(* IEC 61131-3 sources: plc-st-test/packages/core/test/testdata/interpreter, 24 files *)

(* ---- arrays.st ---- *)
(* IEC 61131-3 §6.4.4.4 / Table 15 (ARRAY): bounds are declared as [lo..hi] and may be negative or non-zero based; an element outside the declared bounds is a runtime error; arrays have value semantics on assignment (a copy, not an alias); multi-dimensional arrays index per dimension. *)
FUNCTION_BLOCK TEST_Arrays
VAR
  a : ARRAY[1..5] OF DINT;
  neg : ARRAY[-2..2] OF INT;
  m : ARRAY[0..1, 0..2] OF DINT;
  b : ARRAY[1..5] OF DINT;
  i, idx : DINT;
END_VAR
METHOD Test_FirstAndLastElement
  a[1] := 10;
  a[5] := 50;
  ASSERT_EQUAL_DINT(a[1], 10);
  ASSERT_EQUAL_DINT(a[5], 50);
  ASSERT_EQUAL_DINT(a[3], 0);
END_METHOD
METHOD Test_NegativeLowerBound
  neg[-2] := -20;
  neg[0] := 5;
  neg[2] := 22;
  ASSERT_EQUAL_INT(neg[-2], -20);
  ASSERT_EQUAL_INT(neg[0], 5);
  ASSERT_EQUAL_INT(neg[2], 22);
END_METHOD
METHOD Test_IndexBelowLowerBoundErrors
  idx := 0;
  a[idx] := 1;
END_METHOD
METHOD Test_IndexAboveUpperBoundErrors
  idx := 6;
  i := a[idx];
END_METHOD
METHOD Test_TwoDimensional
  FOR i := 0 TO 2 DO
    m[0, i] := i;
    m[1, i] := 10 + i;
  END_FOR
  ASSERT_EQUAL_DINT(m[0, 2], 2);
  ASSERT_EQUAL_DINT(m[1, 0], 10);
  ASSERT_EQUAL_DINT(m[1, 2], 12);
END_METHOD
METHOD Test_AssignmentCopiesValue
  a[1] := 1; a[2] := 2;
  b := a;
  a[1] := 99;
  ASSERT_EQUAL_DINT(b[1], 1);
  ASSERT_EQUAL_DINT(b[2], 2);
  ASSERT_EQUAL_DINT(a[1], 99);
END_METHOD
METHOD Test_ComputedIndex
  FOR i := 1 TO 5 DO
    a[i] := i * i;
  END_FOR
  ASSERT_EQUAL_DINT(a[a[2]], 16);
END_METHOD
END_FUNCTION_BLOCK

(* ---- bit-operations.st ---- *)
(* IEC 61131-3 §6.6.1 / Table 30 and Table 33: AND/OR/XOR/NOT on bit-string types work bitwise within the type's width (NOT BYTE#16#0F is 16#F0, not a wider value), and BOOL operands use plain logic. *)
FUNCTION_BLOCK TEST_BitOperations
VAR b : BYTE; w : WORD; dw : DWORD; lw : LWORD; END_VAR
METHOD Test_NotStaysInWidth
  b := 16#0F;
  ASSERT_EQUAL_BYTE(NOT b, 16#F0);
  w := 16#00FF;
  ASSERT_EQUAL_WORD(NOT w, 16#FF00);
  dw := 0;
  ASSERT_EQUAL_DWORD(NOT dw, 16#FFFFFFFF);
END_METHOD
METHOD Test_AndOrXor
  b := 16#CC;
  ASSERT_EQUAL_BYTE(b AND 16#0F, 16#0C);
  ASSERT_EQUAL_BYTE(b OR 16#0F, 16#CF);
  ASSERT_EQUAL_BYTE(b XOR 16#FF, 16#33);
END_METHOD
METHOD Test_WordMasks
  w := 16#ABCD;
  ASSERT_EQUAL_WORD(w AND 16#FF00, 16#AB00);
  ASSERT_EQUAL_WORD(w AND 16#00FF, 16#00CD);
  ASSERT_EQUAL_WORD(w XOR w, 0);
END_METHOD
METHOD Test_Lword64BitOps
  lw := 16#8000_0000_0000_0001;
  ASSERT_EQUAL_LWORD(lw AND 16#FFFF_FFFF_0000_0000, 16#8000_0000_0000_0000);
  ASSERT_EQUAL_LWORD(lw OR 16#2, 16#8000_0000_0000_0003);
  ASSERT_EQUAL_LWORD(NOT lw, 16#7FFF_FFFF_FFFF_FFFE);
END_METHOD
METHOD Test_BoolLogicTruthTables
  ASSERT_TRUE(TRUE AND TRUE);
  ASSERT_FALSE(TRUE AND FALSE);
  ASSERT_TRUE(FALSE OR TRUE);
  ASSERT_FALSE(FALSE OR FALSE);
  ASSERT_FALSE(TRUE XOR TRUE);
  ASSERT_TRUE(TRUE XOR FALSE);
  ASSERT_TRUE(NOT FALSE);
  ASSERT_FALSE(NOT TRUE);
END_METHOD
END_FUNCTION_BLOCK

(* ---- case-statement.st ---- *)
(* IEC 61131-3 §6.6.2.5.3 / Table 72 (CASE): selector arms may be single values, comma lists and ranges a..b; ELSE runs when no arm matches; at most one arm runs; enumerated selectors use enumerator labels. *)
TYPE E_Mode : (Off, Manual, Auto, Fault); END_TYPE

FUNCTION_BLOCK TEST_Case
VAR n, r : DINT; m : E_Mode; END_VAR
METHOD Classify
  CASE n OF
    1: r := 10;
    2, 3, 5: r := 20;
    10..19: r := 30;
    -5..-1: r := 40;
  ELSE
    r := 99;
  END_CASE
END_METHOD
METHOD Test_SingleValue
  n := 1; Classify();
  ASSERT_EQUAL_DINT(r, 10);
END_METHOD
METHOD Test_List
  n := 2; Classify();
  ASSERT_EQUAL_DINT(r, 20);
  n := 3; Classify();
  ASSERT_EQUAL_DINT(r, 20);
  n := 5; Classify();
  ASSERT_EQUAL_DINT(r, 20);
END_METHOD
METHOD Test_ListGapFallsToElse
  n := 4; Classify();
  ASSERT_EQUAL_DINT(r, 99);
END_METHOD
METHOD Test_RangeBounds
  n := 10; Classify();
  ASSERT_EQUAL_DINT(r, 30);
  n := 15; Classify();
  ASSERT_EQUAL_DINT(r, 30);
  n := 19; Classify();
  ASSERT_EQUAL_DINT(r, 30);
  n := 9; Classify();
  ASSERT_EQUAL_DINT(r, 99);
  n := 20; Classify();
  ASSERT_EQUAL_DINT(r, 99);
END_METHOD
METHOD Test_NegativeRange
  n := -3; Classify();
  ASSERT_EQUAL_DINT(r, 40);
  n := 0; Classify();
  ASSERT_EQUAL_DINT(r, 99);
END_METHOD
METHOD Test_NoElseNoMatchLeavesUnchanged
  r := 7; n := 50;
  CASE n OF
    1: r := 1;
  END_CASE
  ASSERT_EQUAL_DINT(r, 7);
END_METHOD
METHOD Test_EnumArms
  m := E_Mode.Auto;
  CASE m OF
    E_Mode.Off: r := 0;
    E_Mode.Manual, E_Mode.Auto: r := 1;
    E_Mode.Fault: r := 2;
  END_CASE
  ASSERT_EQUAL_DINT(r, 1);
  m := E_Mode.Fault;
  CASE m OF
    E_Mode.Off: r := 0;
    E_Mode.Manual, E_Mode.Auto: r := 1;
    E_Mode.Fault: r := 2;
  END_CASE
  ASSERT_EQUAL_DINT(r, 2);
END_METHOD
METHOD Test_EnumElse
  m := E_Mode.Manual;
  CASE m OF
    E_Mode.Off: r := 0;
  ELSE
    r := -1;
  END_CASE
  ASSERT_EQUAL_DINT(r, -1);
END_METHOD
METHOD Test_OnlyFirstMatchingArmRuns
  n := 2; r := 0;
  CASE n OF
    1..5: r := r + 1;
    2: r := r + 100;
  END_CASE
  ASSERT_EQUAL_DINT(r, 1);
END_METHOD
END_FUNCTION_BLOCK

(* ---- conversions.st ---- *)
(* IEC 61131-3 §6.6.1 Table 30 note on conversion: REAL/LREAL to an integer type rounds to nearest, ties to even (so 0.5 -> 0, 1.5 -> 2, 2.5 -> 2, -0.5 -> 0, -1.5 -> -2); integer narrowing keeps the low-order bits (two's complement wrap); BOOL converts to 0/1. *)
FUNCTION_BLOCK TEST_Conversions
VAR r : REAL; l : LREAL; i : INT; d : DINT; END_VAR
METHOD Test_RealToIntTiesToEven
  r := 0.5;
  ASSERT_EQUAL_DINT(REAL_TO_DINT(r), 0);
  r := 1.5;
  ASSERT_EQUAL_DINT(REAL_TO_DINT(r), 2);
  r := 2.5;
  ASSERT_EQUAL_DINT(REAL_TO_DINT(r), 2);
  r := 3.5;
  ASSERT_EQUAL_DINT(REAL_TO_DINT(r), 4);
END_METHOD
METHOD Test_NegativeTiesToEven
  r := -0.5;
  ASSERT_EQUAL_DINT(REAL_TO_DINT(r), 0);
  r := -1.5;
  ASSERT_EQUAL_DINT(REAL_TO_DINT(r), -2);
  r := -2.5;
  ASSERT_EQUAL_DINT(REAL_TO_DINT(r), -2);
END_METHOD
METHOD Test_NonTiesRoundToNearest
  l := 2.4;
  ASSERT_EQUAL_DINT(LREAL_TO_DINT(l), 2);
  l := 2.6;
  ASSERT_EQUAL_DINT(LREAL_TO_DINT(l), 3);
  l := -2.6;
  ASSERT_EQUAL_DINT(LREAL_TO_DINT(l), -3);
END_METHOD
METHOD Test_IntNarrowingWraps
  d := 300;
  ASSERT_EQUAL_SINT(DINT_TO_SINT(d), 44);
  d := 70000;
  ASSERT_EQUAL_INT(DINT_TO_INT(d), 4464);
  d := -1;
  ASSERT_EQUAL_USINT(DINT_TO_USINT(d), 255);
END_METHOD
METHOD Test_WideningPreservesValue
  i := -5;
  ASSERT_EQUAL_DINT(INT_TO_DINT(i), -5);
  ASSERT_EQUAL_LINT(INT_TO_LINT(i), -5);
  ASSERT_EQUAL_REAL(INT_TO_REAL(i), -5.0);
END_METHOD
METHOD Test_BoolConversions
  ASSERT_EQUAL_DINT(BOOL_TO_DINT(TRUE), 1);
  ASSERT_EQUAL_DINT(BOOL_TO_DINT(FALSE), 0);
  d := 7;
  ASSERT_TRUE(DINT_TO_BOOL(d));
  d := 0;
  ASSERT_FALSE(DINT_TO_BOOL(d));
END_METHOD
METHOD Test_UnsignedFromNegativeWraps
  d := -1;
  ASSERT_EQUAL_UDINT(DINT_TO_UDINT(d), 4294967295);
END_METHOD
END_FUNCTION_BLOCK

(* ---- counters-edges.st ---- *)
(* IEC 61131-3 §6.6.3.2 / Tables 41-42 (CTU, CTD) and R_TRIG/F_TRIG (Table 40): counters count only on a rising edge of CU/CD evaluated once per cycle, so holding the input TRUE for many cycles counts once; CTU.Q = (CV >= PV); R_TRIG.Q is TRUE for exactly the cycle in which CLK rose. *)
FUNCTION_BLOCK TEST_CountersEdges
VAR
  ctu : CTU;
  rt : R_TRIG;
  ft : F_TRIG;
  clk : BOOL;
  rst : BOOL;
  rises, falls : DINT;
END_VAR
METHOD Cycle
  ctu(CU := clk, R := rst, PV := 3);
  rt(CLK := clk);
  ft(CLK := clk);
  IF rt.Q THEN rises := rises + 1; END_IF
  IF ft.Q THEN falls := falls + 1; END_IF
END_METHOD
METHOD Test_HeldInputCountsOnce
  clk := TRUE;
  RUN_CYCLES(10);
  ASSERT_EQUAL_INT(ctu.CV, 1);
  ASSERT_EQUAL_DINT(rises, 1);
  ASSERT_EQUAL_DINT(falls, 0);
END_METHOD
METHOD Test_ToggleCountsEachRisingEdge
  clk := TRUE;  RUN_CYCLES(1);
  clk := FALSE; RUN_CYCLES(1);
  clk := TRUE;  RUN_CYCLES(1);
  clk := FALSE; RUN_CYCLES(1);
  ASSERT_EQUAL_INT(ctu.CV, 2);
  ASSERT_EQUAL_DINT(rises, 2);
  ASSERT_EQUAL_DINT(falls, 2);
  ASSERT_FALSE(ctu.Q);
END_METHOD
METHOD Test_QSetsAtPreset
  clk := TRUE;  RUN_CYCLES(1);
  clk := FALSE; RUN_CYCLES(1);
  clk := TRUE;  RUN_CYCLES(1);
  clk := FALSE; RUN_CYCLES(1);
  clk := TRUE;  RUN_CYCLES(1);
  ASSERT_EQUAL_INT(ctu.CV, 3);
  ASSERT_TRUE(ctu.Q);
END_METHOD
METHOD Test_ResetClearsCountAndQ
  clk := TRUE;  RUN_CYCLES(1);
  clk := FALSE; RUN_CYCLES(1);
  clk := TRUE;  RUN_CYCLES(1);
  clk := FALSE; RUN_CYCLES(1);
  clk := TRUE;  RUN_CYCLES(1);
  rst := TRUE;
  RUN_CYCLES(1);
  ASSERT_EQUAL_INT(ctu.CV, 0);
  ASSERT_FALSE(ctu.Q);
END_METHOD
METHOD Test_PulseOnlyOneCycleWide
  clk := TRUE;
  RUN_CYCLES(1);
  ASSERT_TRUE(rt.Q);
  RUN_CYCLES(1);
  ASSERT_FALSE(rt.Q);
END_METHOD
END_FUNCTION_BLOCK

(* ---- deep-nesting.st ---- *)
(* IEC 61131-3 §6.6.2 (statements compose freely): IF/ELSIF/ELSE, CASE and loops nest to arbitrary depth with the innermost branch selected by the combined conditions; expressions nest through parentheses with the Table 71 precedence (NOT, **, unary minus, * / MOD, + -, comparisons, AND, XOR, OR). *)
FUNCTION_BLOCK TEST_DeepNesting
VAR a, b, c, r, i, j, k, count : DINT; ok : BOOL; END_VAR
METHOD Test_NestedIfElsifChain
  a := 2; b := 3; c := 4;
  IF a = 1 THEN
    r := 1;
  ELSIF a = 2 THEN
    IF b = 2 THEN
      r := 2;
    ELSIF b = 3 THEN
      IF c = 3 THEN
        r := 3;
      ELSE
        IF c = 4 THEN r := 4; ELSE r := 5; END_IF
      END_IF
    END_IF
  ELSE
    r := 6;
  END_IF
  ASSERT_EQUAL_DINT(r, 4);
END_METHOD
METHOD Test_TripleNestedLoopCount
  count := 0;
  FOR i := 1 TO 4 DO
    FOR j := 1 TO 3 DO
      FOR k := 1 TO 2 DO
        count := count + 1;
      END_FOR
    END_FOR
  END_FOR
  ASSERT_EQUAL_DINT(count, 24);
END_METHOD
METHOD Test_LoopsCaseAndIfTogether
  count := 0;
  FOR i := 1 TO 6 DO
    CASE i MOD 3 OF
      0: count := count + 100;
      1:
        IF i > 3 THEN count := count + 10; ELSE count := count + 1; END_IF
    ELSE
      count := count + 1000;
    END_CASE
  END_FOR
  ASSERT_EQUAL_DINT(count, 2 * 1000 + 2 * 100 + 10 + 1);
END_METHOD
METHOD Test_ParenthesesNestDeeply
  a := 2;
  r := ((((a + 1) * (a + 2)) - ((a - 1) * (a + 3))) * 2) + (((a)));
  ASSERT_EQUAL_DINT(r, 16);
END_METHOD
METHOD Test_PrecedenceTable71
  r := 2 + 3 * 4;
  ASSERT_EQUAL_DINT(r, 14);
  r := 20 - 6 / 3 - 1;
  ASSERT_EQUAL_DINT(r, 17);
  r := 2 * 3 MOD 4;
  ASSERT_EQUAL_DINT(r, 2);
  r := -2 * 3;
  ASSERT_EQUAL_DINT(r, -6);
END_METHOD
METHOD Test_BooleanPrecedence
  ok := TRUE OR FALSE AND FALSE;
  ASSERT_TRUE(ok);
  ok := NOT FALSE AND FALSE;
  ASSERT_FALSE(ok);
  ok := TRUE XOR TRUE OR TRUE;
  ASSERT_TRUE(ok);
  a := 1; b := 2;
  ok := a < b AND b < 3 OR FALSE;
  ASSERT_TRUE(ok);
END_METHOD
METHOD Test_WhileInsideRepeatInsideFor
  count := 0;
  FOR i := 1 TO 2 DO
    j := 0;
    REPEAT
      j := j + 1;
      k := 0;
      WHILE k < 2 DO
        k := k + 1;
        count := count + 1;
      END_WHILE
    UNTIL j >= 3
    END_REPEAT
  END_FOR
  ASSERT_EQUAL_DINT(count, 12);
END_METHOD
END_FUNCTION_BLOCK

(* ---- division.st ---- *)
(* IEC 61131-3 §6.6.1.4 / Table 30: division by zero is an error for integer and real operands, and for MOD; this runtime raises IecRuntimeError 'division by zero' (test errored). Also integer division truncates toward zero. *)
FUNCTION_BLOCK TEST_Division
VAR i, z : DINT; r, rz : REAL; l, lz : LREAL; END_VAR
METHOD Test_IntDivByZeroErrors
  z := 0; i := 5 / z;
END_METHOD
METHOD Test_RealDivByZeroErrors
  rz := 0.0; r := 1.0 / rz;
END_METHOD
METHOD Test_LrealDivByZeroErrors
  lz := 0.0; l := 1.0 / lz;
END_METHOD
METHOD Test_ModByZeroErrors
  z := 0; i := 5 MOD z;
END_METHOD
METHOD Test_IntDivTruncatesTowardZero
  i := 7; z := 2;
  ASSERT_EQUAL_DINT(i / z, 3);
  i := -7;
  ASSERT_EQUAL_DINT(i / z, -3);
  z := -2;
  ASSERT_EQUAL_DINT(i / z, 3);
  i := 7;
  ASSERT_EQUAL_DINT(i / z, -3);
END_METHOD
METHOD Test_RealDivNormal
  r := 1.0; rz := 4.0;
  ASSERT_EQUAL_REAL(r / rz, 0.25);
END_METHOD
END_FUNCTION_BLOCK

(* ---- enums.st ---- *)
(* IEC 61131-3 §6.4.4.2 / Table 12 (enumerated data types): enumerators without an explicit value number from 0 and continue from the previous value after an explicit one; a variable of enumerated type starts at its first enumerator unless an initial value is given; enumerators of one type compare by value. *)
TYPE E_Color : (Red, Green := 5, Blue); END_TYPE
TYPE E_Level : (Low, Mid, High) := Mid; END_TYPE

FUNCTION_BLOCK TEST_Enums
VAR
  c : E_Color;
  lv : E_Level;
  c2 : E_Color := E_Color.Blue;
  n : DINT;
END_VAR
METHOD Test_DefaultIsFirstEnumerator
  ASSERT_EQUAL(c, E_Color.Red);
END_METHOD
METHOD Test_DeclaredInitialValue
  ASSERT_EQUAL(c2, E_Color.Blue);
END_METHOD
METHOD Test_TypeLevelDefault
  ASSERT_EQUAL(lv, E_Level.Mid);
END_METHOD
METHOD Test_ExplicitAndImplicitValues
  n := E_Color.Red;
  ASSERT_EQUAL_DINT(n, 0);
  n := E_Color.Green;
  ASSERT_EQUAL_DINT(n, 5);
  n := E_Color.Blue;
  ASSERT_EQUAL_DINT(n, 6);
END_METHOD
METHOD Test_Comparison
  c := E_Color.Green;
  ASSERT_TRUE(c = E_Color.Green);
  ASSERT_TRUE(c <> E_Color.Blue);
  ASSERT_NOT_EQUAL(c, E_Color.Red);
END_METHOD
METHOD Test_AssignAndCopy
  c := E_Color.Blue;
  c2 := c;
  c := E_Color.Red;
  ASSERT_EQUAL(c2, E_Color.Blue);
  ASSERT_EQUAL(c, E_Color.Red);
END_METHOD
END_FUNCTION_BLOCK

(* ---- fb-instances.st ---- *)
(* IEC 61131-3 §6.6.3 (function blocks): every FB instance has its own copy of the internal VAR state, instances do not share data, and state persists between calls of the same instance. Struct assignment (§6.4.4.3) copies all members. *)
TYPE ST_Point : STRUCT x : DINT; y : DINT; END_STRUCT; END_TYPE

FUNCTION_BLOCK FB_Acc
VAR_INPUT step : DINT; END_VAR
VAR total : DINT; END_VAR
VAR_OUTPUT out : DINT; END_VAR
METHOD Add
  total := total + step;
  out := total;
END_METHOD
END_FUNCTION_BLOCK

FUNCTION_BLOCK TEST_FbInstances
VAR
  a, b : FB_Acc;
  p, q : ST_Point;
  r : DINT;
END_VAR
METHOD Test_InstancesAreIndependent
  a.step := 1; b.step := 10;
  a.Add(); a.Add(); b.Add();
  ASSERT_EQUAL_DINT(a.total, 2);
  ASSERT_EQUAL_DINT(b.total, 10);
END_METHOD
METHOD Test_StatePersistsBetweenCalls
  a.step := 5;
  a.Add(); a.Add(); a.Add();
  ASSERT_EQUAL_DINT(a.out, 15);
END_METHOD
METHOD Test_OutputReadAfterCall
  b.step := 3;
  b.Add();
  r := b.out;
  ASSERT_EQUAL_DINT(r, 3);
END_METHOD
METHOD Test_StructAssignmentCopies
  p.x := 1; p.y := 2;
  q := p;
  p.x := 100;
  ASSERT_EQUAL_DINT(q.x, 1);
  ASSERT_EQUAL_DINT(q.y, 2);
  ASSERT_EQUAL_DINT(p.x, 100);
END_METHOD
METHOD Test_FreshInstanceHasZeroState
  ASSERT_EQUAL_DINT(a.total, 0);
  ASSERT_EQUAL_DINT(p.x, 0);
END_METHOD
END_FUNCTION_BLOCK

(* ---- for-loops.st ---- *)
(* IEC 61131-3 §6.6.2.5.4 / Table 72 (FOR): the body runs while the control variable has not passed the end value in the direction of BY; a negative BY counts down; when start already passes end the body runs zero times. *)
FUNCTION_BLOCK TEST_ForLoops
VAR i, n, sum : DINT; END_VAR
METHOD Test_NegativeStep
  sum := 0; n := 0;
  FOR i := 10 TO 1 BY -3 DO
    sum := sum + i;
    n := n + 1;
  END_FOR
  ASSERT_EQUAL_DINT(sum, 22);
  ASSERT_EQUAL_DINT(n, 4);
END_METHOD
METHOD Test_ZeroIterations
  n := 0;
  FOR i := 5 TO 4 DO
    n := n + 1;
  END_FOR
  ASSERT_EQUAL_DINT(n, 0);
END_METHOD
METHOD Test_ZeroIterationsNegativeStep
  n := 0;
  FOR i := 1 TO 5 BY -1 DO
    n := n + 1;
  END_FOR
  ASSERT_EQUAL_DINT(n, 0);
END_METHOD
METHOD Test_SingleIteration
  n := 0;
  FOR i := 3 TO 3 DO
    n := n + 1;
  END_FOR
  ASSERT_EQUAL_DINT(n, 1);
END_METHOD
METHOD Test_DefaultStepOne
  sum := 0;
  FOR i := 1 TO 5 DO
    sum := sum + i;
  END_FOR
  ASSERT_EQUAL_DINT(sum, 15);
END_METHOD
METHOD Test_PositiveStepTwo
  sum := 0;
  FOR i := 0 TO 10 BY 2 DO
    sum := sum + i;
  END_FOR
  ASSERT_EQUAL_DINT(sum, 30);
END_METHOD
METHOD Test_LastValueSeenInBody
  FOR i := 1 TO 3 DO
    n := i;
  END_FOR
  ASSERT_EQUAL_DINT(n, 3);
END_METHOD
METHOD Test_NegativeRange
  sum := 0;
  FOR i := -2 TO 2 DO
    sum := sum + i * i;
  END_FOR
  ASSERT_EQUAL_DINT(sum, 10);
END_METHOD
END_FUNCTION_BLOCK

(* ---- initial-values.st ---- *)
(* IEC 61131-3 §6.4.2 / Table 62 (default initial values): every variable without an explicit initializer starts at the type's default (0, FALSE, empty string, T#0s, first enumerator); explicit initializers, including constant expressions and negative literals, override it; FB instances start fresh for every test. *)
FUNCTION_BLOCK TEST_InitialValues
VAR CONSTANT
  K : DINT := 4;
END_VAR
VAR
  i : INT;
  u : UDINT;
  r : REAL;
  b : BOOL;
  s : STRING;
  t : TIME;
  l : LINT;
  neg : INT := -7;
  expr : DINT := K * 2 + 1;
  arr : ARRAY[0..2] OF DINT := [1, 2, 3];
  zeros : ARRAY[0..2] OF BYTE;
END_VAR
METHOD Test_NumericDefaultsAreZero
  ASSERT_EQUAL_INT(i, 0);
  ASSERT_EQUAL_UDINT(u, 0);
  ASSERT_EQUAL_REAL(r, 0.0);
  ASSERT_EQUAL_LINT(l, 0);
END_METHOD
METHOD Test_BoolStringTimeDefaults
  ASSERT_FALSE(b);
  ASSERT_EQUAL_STRING(s, '');
  ASSERT_EQUAL_TIME(t, T#0s);
END_METHOD
METHOD Test_NegativeInitializer
  ASSERT_EQUAL_INT(neg, -7);
END_METHOD
METHOD Test_ConstantExpressionInitializer
  ASSERT_EQUAL_DINT(expr, 9);
END_METHOD
METHOD Test_ArrayInitializer
  ASSERT_EQUAL_DINT(arr[0], 1);
  ASSERT_EQUAL_DINT(arr[2], 3);
  ASSERT_EQUAL_BYTE(zeros[1], 0);
END_METHOD
METHOD Test_StateDoesNotLeakBetweenTests
  i := 42;
  s := 'dirty';
END_METHOD
METHOD Test_FreshAfterDirtyingTest
  ASSERT_EQUAL_INT(i, 0);
  ASSERT_EQUAL_STRING(s, '');
END_METHOD
END_FUNCTION_BLOCK

(* ---- loop-exit-continue.st ---- *)
(* IEC 61131-3 §6.6.2.5.4 (EXIT) and ed.3 CONTINUE: EXIT leaves only the innermost enclosing loop; CONTINUE skips to the next iteration of the innermost loop. Applies to FOR, WHILE and REPEAT. *)
FUNCTION_BLOCK TEST_LoopExitContinue
VAR i, j, n, outer, inner : DINT; END_VAR
METHOD Test_ExitLeavesInnermostOnly
  outer := 0; inner := 0;
  FOR i := 1 TO 3 DO
    outer := outer + 1;
    FOR j := 1 TO 10 DO
      IF j = 3 THEN EXIT; END_IF
      inner := inner + 1;
    END_FOR
  END_FOR
  ASSERT_EQUAL_DINT(outer, 3);
  ASSERT_EQUAL_DINT(inner, 6);
END_METHOD
METHOD Test_ContinueSkipsRestOfBody
  n := 0;
  FOR i := 1 TO 5 DO
    IF i MOD 2 = 0 THEN CONTINUE; END_IF
    n := n + i;
  END_FOR
  ASSERT_EQUAL_DINT(n, 9);
END_METHOD
METHOD Test_ContinueInInnerOnly
  outer := 0; inner := 0;
  FOR i := 1 TO 2 DO
    outer := outer + 1;
    FOR j := 1 TO 4 DO
      IF j <= 2 THEN CONTINUE; END_IF
      inner := inner + 1;
    END_FOR
  END_FOR
  ASSERT_EQUAL_DINT(outer, 2);
  ASSERT_EQUAL_DINT(inner, 4);
END_METHOD
METHOD Test_ExitFromWhile
  n := 0;
  WHILE TRUE DO
    n := n + 1;
    IF n = 7 THEN EXIT; END_IF
  END_WHILE
  ASSERT_EQUAL_DINT(n, 7);
END_METHOD
METHOD Test_ExitFromRepeat
  n := 0;
  REPEAT
    n := n + 1;
    IF n = 4 THEN EXIT; END_IF
  UNTIL FALSE
  END_REPEAT
  ASSERT_EQUAL_DINT(n, 4);
END_METHOD
METHOD Test_ContinueInRepeatStillEvaluatesUntil
  n := 0; i := 0;
  REPEAT
    i := i + 1;
    IF i < 3 THEN CONTINUE; END_IF
    n := n + 1;
  UNTIL i >= 5
  END_REPEAT
  ASSERT_EQUAL_DINT(n, 3);
  ASSERT_EQUAL_DINT(i, 5);
END_METHOD
METHOD Test_ExitInMixedNesting
  n := 0;
  FOR i := 1 TO 3 DO
    j := 0;
    WHILE TRUE DO
      j := j + 1;
      IF j > 2 THEN EXIT; END_IF
      n := n + 1;
    END_WHILE
  END_FOR
  ASSERT_EQUAL_DINT(n, 6);
END_METHOD
METHOD Test_WhileZeroIterations
  n := 0;
  WHILE FALSE DO n := 1; END_WHILE
  ASSERT_EQUAL_DINT(n, 0);
END_METHOD
METHOD Test_RepeatRunsAtLeastOnce
  n := 0;
  REPEAT n := n + 1; UNTIL TRUE END_REPEAT
  ASSERT_EQUAL_DINT(n, 1);
END_METHOD
END_FUNCTION_BLOCK

(* ---- mod-negative.st ---- *)
(* IEC 61131-3 §6.6.1.4 Table 30 (MOD): IN1 MOD IN2 = IN1 - (IN1/IN2)*IN2 with truncating division, so the result takes the sign of the dividend. *)
FUNCTION_BLOCK TEST_ModNegative
VAR a, b : DINT; la, lb : LINT; END_VAR
METHOD Test_PositivePositive
  a := 7; b := 3;
  ASSERT_EQUAL_DINT(a MOD b, 1);
END_METHOD
METHOD Test_NegativeDividend
  a := -7; b := 3;
  ASSERT_EQUAL_DINT(a MOD b, -1);
END_METHOD
METHOD Test_NegativeDivisor
  a := 7; b := -3;
  ASSERT_EQUAL_DINT(a MOD b, 1);
END_METHOD
METHOD Test_BothNegative
  a := -7; b := -3;
  ASSERT_EQUAL_DINT(a MOD b, -1);
END_METHOD
METHOD Test_ExactMultipleIsZero
  a := -9; b := 3;
  ASSERT_EQUAL_DINT(a MOD b, 0);
END_METHOD
METHOD Test_BigIntNegative
  la := -7; lb := 3;
  ASSERT_EQUAL_LINT(la MOD lb, -1);
  la := 7; lb := -3;
  ASSERT_EQUAL_LINT(la MOD lb, 1);
END_METHOD
END_FUNCTION_BLOCK

(* ---- overflow-bigint.st ---- *)
(* IEC 61131-3 §6.6.1 / Table 30: 64-bit types wrap modulo 2^64: LINT -2^63..2^63-1, ULINT 0..2^64-1, LWORD 0..2^64-1 (bit string). Values beyond 2^53 must stay exact. *)
FUNCTION_BLOCK TEST_OverflowBigint
VAR l : LINT; ul : ULINT; lw : LWORD; END_VAR
METHOD Test_LintPositiveWrap
  l := 9223372036854775807; l := l + 1;
  ASSERT_EQUAL_LINT(l, -9223372036854775808);
END_METHOD
METHOD Test_LintNegativeWrap
  l := -9223372036854775808; l := l - 1;
  ASSERT_EQUAL_LINT(l, 9223372036854775807);
END_METHOD
METHOD Test_UlintWrap
  ul := 18446744073709551615; ul := ul + 1;
  ASSERT_EQUAL_ULINT(ul, 0);
  ul := 0; ul := ul - 1;
  ASSERT_EQUAL_ULINT(ul, 18446744073709551615);
END_METHOD
METHOD Test_LwordWrap
  lw := 16#FFFF_FFFF_FFFF_FFFF; lw := lw + 1;
  ASSERT_EQUAL_LWORD(lw, 0);
END_METHOD
METHOD Test_PrecisionBeyond2Pow53
  l := 9007199254740993;
  ASSERT_EQUAL_LINT(l, 9007199254740993);
  l := l + 1;
  ASSERT_EQUAL_LINT(l, 9007199254740994);
END_METHOD
METHOD Test_LintMultiplyWrap
  l := 4294967296; l := l * 4294967296;
  ASSERT_EQUAL_LINT(l, 0);
END_METHOD
END_FUNCTION_BLOCK

(* ---- overflow-dint.st ---- *)
(* IEC 61131-3 §6.6.1 / Table 30: DINT (-2^31..2^31-1) and UDINT (0..2^32-1) arithmetic wraps modulo 2^32. *)
FUNCTION_BLOCK TEST_OverflowDint
VAR d : DINT; ud : UDINT; END_VAR
METHOD Test_DintPositiveWrap
  d := 2147483647; d := d + 1;
  ASSERT_EQUAL_DINT(d, -2147483648);
END_METHOD
METHOD Test_DintNegativeWrap
  d := -2147483648; d := d - 1;
  ASSERT_EQUAL_DINT(d, 2147483647);
END_METHOD
METHOD Test_UdintWrap
  ud := 4294967295; ud := ud + 1;
  ASSERT_EQUAL_UDINT(ud, 0);
  ud := 0; ud := ud - 1;
  ASSERT_EQUAL_UDINT(ud, 4294967295);
END_METHOD
METHOD Test_DintMultiplyWrap
  d := 65536; d := d * 65536;
  ASSERT_EQUAL_DINT(d, 0);
  d := 65537; d := d * 65537;
  ASSERT_EQUAL_DINT(d, 131073);
END_METHOD
METHOD Test_UdintMultiplyWrap
  ud := 4294967295; ud := ud * 2;
  ASSERT_EQUAL_UDINT(ud, 4294967294);
END_METHOD
END_FUNCTION_BLOCK

(* ---- overflow-small-ints.st ---- *)
(* IEC 61131-3 §6.6.1 / Table 30: integer arithmetic on a fixed-width type wraps modulo 2^N on assignment (two's complement): SINT -128..127, USINT 0..255, INT -32768..32767, UINT 0..65535. *)
FUNCTION_BLOCK TEST_OverflowSmall
VAR s : SINT; us : USINT; i : INT; ui : UINT; END_VAR
METHOD Test_SintPositiveWrap
  s := 127; s := s + 1;
  ASSERT_EQUAL_SINT(s, -128);
END_METHOD
METHOD Test_SintNegativeWrap
  s := -128; s := s - 1;
  ASSERT_EQUAL_SINT(s, 127);
END_METHOD
METHOD Test_UsintWrap
  us := 255; us := us + 1;
  ASSERT_EQUAL_USINT(us, 0);
  us := 0; us := us - 1;
  ASSERT_EQUAL_USINT(us, 255);
END_METHOD
METHOD Test_IntWrap
  i := 32767; i := i + 1;
  ASSERT_EQUAL_INT(i, -32768);
  i := -32768; i := i - 1;
  ASSERT_EQUAL_INT(i, 32767);
END_METHOD
METHOD Test_UintWrap
  ui := 65535; ui := ui + 1;
  ASSERT_EQUAL_UINT(ui, 0);
  ui := 0; ui := ui - 1;
  ASSERT_EQUAL_UINT(ui, 65535);
END_METHOD
METHOD Test_MultiplyWrap
  s := 100; s := s * 2;
  ASSERT_EQUAL_SINT(s, -56);
  us := 200; us := us * 2;
  ASSERT_EQUAL_USINT(us, 144);
END_METHOD
METHOD Test_NegateMinimum
  s := -128; s := -s;
  ASSERT_EQUAL_SINT(s, -128);
END_METHOD
END_FUNCTION_BLOCK

(* ---- real-fround.st ---- *)
(* IEC 61131-3 §6.3.2 / Table 10: REAL is IEEE 754 binary32 and LREAL is binary64, so every REAL result is rounded to single precision. 16777217 (2^24+1) is not representable in binary32 and rounds to 16777216. *)
FUNCTION_BLOCK TEST_RealFround
VAR r, r2 : REAL; l, l2 : LREAL; END_VAR
METHOD Test_SinglePrecisionRoundsInteger
  r := 16777217.0;
  ASSERT_EQUAL_REAL(r, 16777216.0);
END_METHOD
METHOD Test_DoubleKeepsInteger
  l := 16777217.0;
  ASSERT_EQUAL_LREAL(l, 16777217.0);
END_METHOD
METHOD Test_LrealZeroPointOnePlusZeroPointTwo
  l := 0.1; l2 := 0.2;
  ASSERT_NEAR(l + l2, 0.3, 1.0E-15);
  ASSERT_NOT_EQUAL_LREAL(l + l2, 0.3);
END_METHOD
METHOD Test_RealZeroPointOnePlusZeroPointTwo
  r := 0.1; r2 := 0.2;
  ASSERT_EQUAL_REAL(r + r2, 0.3);
END_METHOD
METHOD Test_RealAccumulationAbsorbed
  r := 16777216.0;
  r := r + 1.0;
  ASSERT_EQUAL_REAL(r, 16777216.0);
END_METHOD
METHOD Test_LrealAccumulationKept
  l := 16777216.0;
  l := l + 1.0;
  ASSERT_EQUAL_LREAL(l, 16777217.0);
END_METHOD
METHOD Test_RealStoresRoundedDouble
  l := 0.1;
  r := l;
  l2 := r;
  ASSERT_NOT_EQUAL_LREAL(l2, 0.1);
  ASSERT_NEAR(l2, 0.1, 1.0E-7);
END_METHOD
END_FUNCTION_BLOCK

(* ---- recursion.st ---- *)
(* IEC 61131-3 §6.6.1.5 leaves recursion implementation-defined (the standard does not permit a function to call itself); this runtime allows bounded recursion and ends a runaway one with a limit error (test errored, kind limit) instead of a stack overflow. *)
FUNCTION F_Factorial : DINT
VAR_INPUT n : DINT; END_VAR
IF n <= 1 THEN
  F_Factorial := 1;
ELSE
  F_Factorial := n * F_Factorial(n - 1);
END_IF
END_FUNCTION

FUNCTION F_Runaway : DINT
VAR_INPUT n : DINT; END_VAR
F_Runaway := F_Runaway(n + 1);
END_FUNCTION

FUNCTION F_Depth : DINT
VAR_INPUT n : DINT; END_VAR
IF n = 0 THEN
  F_Depth := 0;
ELSE
  F_Depth := 1 + F_Depth(n - 1);
END_IF
END_FUNCTION

FUNCTION_BLOCK TEST_Recursion
METHOD Test_FactorialShallow
  ASSERT_EQUAL_DINT(F_Factorial(5), 120);
  ASSERT_EQUAL_DINT(F_Factorial(1), 1);
  ASSERT_EQUAL_DINT(F_Factorial(10), 3628800);
END_METHOD
METHOD Test_RunawayRecursionHitsLimit
  ASSERT_EQUAL_DINT(F_Runaway(0), 0);
END_METHOD
METHOD Test_ModerateDepthOk
  ASSERT_EQUAL_DINT(F_Depth(50), 50);
END_METHOD
END_FUNCTION_BLOCK

(* ---- return-method.st ---- *)
(* IEC 61131-3 §6.6.2.4 / Table 72 (RETURN): RETURN ends the current POU invocation immediately; statements after it are not executed, a result assigned before RETURN is the returned value, and only the current method is left, not the caller. *)
FUNCTION_BLOCK FB_Guard
VAR
  calls : DINT;
  reached : DINT;
END_VAR
METHOD Early : DINT
VAR_INPUT x : DINT; END_VAR
  calls := calls + 1;
  Early := 1;
  IF x < 0 THEN
    RETURN;
  END_IF
  reached := reached + 1;
  Early := 2;
END_METHOD
METHOD InLoop : DINT
VAR_INPUT limit : DINT; END_VAR
VAR k : DINT; END_VAR
  FOR k := 1 TO 100 DO
    IF k = limit THEN
      InLoop := k;
      RETURN;
    END_IF
  END_FOR
  InLoop := -1;
END_METHOD
METHOD Inner
  RETURN;
END_METHOD
METHOD Outer : DINT
  Outer := 10;
  Inner();
  Outer := Outer + 1;
END_METHOD
END_FUNCTION_BLOCK

FUNCTION_BLOCK TEST_ReturnMethod
VAR g : FB_Guard; r : DINT; END_VAR
METHOD Test_ReturnSkipsRest
  r := g.Early(-1);
  ASSERT_EQUAL_DINT(r, 1);
  ASSERT_EQUAL_DINT(g.reached, 0);
END_METHOD
METHOD Test_NoReturnRunsToEnd
  r := g.Early(5);
  ASSERT_EQUAL_DINT(r, 2);
  ASSERT_EQUAL_DINT(g.reached, 1);
END_METHOD
METHOD Test_ReturnFromInsideLoop
  r := g.InLoop(7);
  ASSERT_EQUAL_DINT(r, 7);
  r := g.InLoop(1000);
  ASSERT_EQUAL_DINT(r, -1);
END_METHOD
METHOD Test_ReturnDoesNotLeaveCaller
  r := g.Outer();
  ASSERT_EQUAL_DINT(r, 11);
END_METHOD
METHOD Test_ReturnInTestMethodStopsIt
  r := 1;
  RETURN;
  r := 2;
  ASSERT_EQUAL_DINT(r, 1);
END_METHOD
METHOD Test_StateAfterReturn
  r := g.Early(-1);
  r := g.Early(-1);
  ASSERT_EQUAL_DINT(g.calls, 2);
END_METHOD
END_FUNCTION_BLOCK

(* ---- string-truncation.st ---- *)
(* IEC 61131-3 §6.3.3 / Table 10 (STRING[n]): a STRING variable declared with length n holds at most n characters; a longer value assigned to it is truncated on the right. *)
FUNCTION_BLOCK TEST_StringTruncation
VAR s : STRING(5); t : STRING(3); u : STRING(255); END_VAR
METHOD Test_AssignTruncates
  s := 'HELLOWORLD';
  ASSERT_EQUAL_STRING(s, 'HELLO');
  ASSERT_EQUAL_INT(LEN(s), 5);
END_METHOD
METHOD Test_ShorterUnchanged
  s := 'AB';
  ASSERT_EQUAL_STRING(s, 'AB');
  ASSERT_EQUAL_INT(LEN(s), 2);
END_METHOD
METHOD Test_ExactLengthUnchanged
  s := 'ABCDE';
  ASSERT_EQUAL_STRING(s, 'ABCDE');
END_METHOD
METHOD Test_ConcatIntoShortTruncates
  t := CONCAT('AB', 'CDEF');
  ASSERT_EQUAL_STRING(t, 'ABC');
END_METHOD
METHOD Test_ConcatWideKeepsAll
  u := CONCAT('AB', 'CDEF');
  ASSERT_EQUAL_STRING(u, 'ABCDEF');
  ASSERT_EQUAL_INT(LEN(u), 6);
END_METHOD
METHOD Test_CopyBetweenStringsTruncates
  u := 'ABCDEFGH';
  t := u;
  ASSERT_EQUAL_STRING(t, 'ABC');
  ASSERT_EQUAL_STRING(u, 'ABCDEFGH');
END_METHOD
METHOD Test_EmptyString
  s := '';
  ASSERT_EQUAL_INT(LEN(s), 0);
END_METHOD
END_FUNCTION_BLOCK

(* ---- temp-vs-var.st ---- *)
(* IEC 61131-3 §6.5.3 / Table 14: VAR keeps its value between invocations of an FB instance, while VAR_TEMP is re-initialised on every invocation. *)
FUNCTION_BLOCK FB_Counter
VAR
  persistent : DINT := 100;
  lastScratch : DINT;
END_VAR
VAR_TEMP
  scratch : DINT := 7;
END_VAR
METHOD Run
  persistent := persistent + 1;
  scratch := scratch + 10;
  lastScratch := scratch;
END_METHOD
END_FUNCTION_BLOCK

FUNCTION_BLOCK FB_TempOnly
VAR_TEMP
  t : DINT;
END_VAR
VAR
  seenNonZero : BOOL;
END_VAR
METHOD Run
  IF t <> 0 THEN seenNonZero := TRUE; END_IF
  t := t + 5;
END_METHOD
END_FUNCTION_BLOCK

FUNCTION_BLOCK TEST_TempVsVar
VAR
  c : FB_Counter;
  o : FB_TempOnly;
  runs : DINT;
END_VAR
METHOD Cycle
  c.Run();
  o.Run();
  runs := runs + 1;
END_METHOD
METHOD Test_VarPersistsAcrossCycles
  RUN_CYCLES(5);
  ASSERT_EQUAL_DINT(c.persistent, 105);
  ASSERT_EQUAL_DINT(runs, 5);
END_METHOD
METHOD Test_VarTempResetsEachInvocation
  RUN_CYCLES(4);
  ASSERT_FALSE(o.seenNonZero);
END_METHOD
METHOD Test_VarTempReinitialisedToDeclaredValue
  RUN_CYCLES(3);
  ASSERT_EQUAL_DINT(c.lastScratch, 17);
END_METHOD
END_FUNCTION_BLOCK

(* ---- time-arithmetic.st ---- *)
(* IEC 61131-3 §6.3.3 / Table 8-9 (TIME): TIME literals combine units (T#1s500ms = 1500 ms); TIME + TIME, TIME - TIME and TIME * number give TIME; TIME values compare chronologically; TIME has no wraparound at the sizes used here. *)
FUNCTION_BLOCK TEST_TimeArithmetic
VAR a, b : TIME; END_VAR
METHOD Test_CompoundLiteral
  a := T#1s500ms;
  ASSERT_EQUAL_TIME(a, T#1500ms);
END_METHOD
METHOD Test_Addition
  a := T#2s; b := T#750ms;
  ASSERT_EQUAL_TIME(a + b, T#2750ms);
END_METHOD
METHOD Test_Subtraction
  a := T#2s; b := T#750ms;
  ASSERT_EQUAL_TIME(a - b, T#1250ms);
END_METHOD
METHOD Test_Comparison
  a := T#1m; b := T#59s;
  ASSERT_TRUE(a > b);
  ASSERT_TRUE(b < a);
  ASSERT_TRUE(a >= T#60s);
  ASSERT_TRUE(a = T#60s);
  ASSERT_TRUE(a <> b);
END_METHOD
METHOD Test_UnitConversions
  ASSERT_EQUAL_TIME(T#1h, T#60m);
  ASSERT_EQUAL_TIME(T#1d, T#24h);
  ASSERT_EQUAL_TIME(T#1s, T#1000ms);
  ASSERT_EQUAL_TIME(T#1ms, T#1000us);
END_METHOD
METHOD Test_ZeroTime
  a := T#0s;
  ASSERT_EQUAL_TIME(a, T#0ms);
  ASSERT_EQUAL_TIME(a + T#5ms, T#5ms);
END_METHOD
END_FUNCTION_BLOCK

(* ---- timers-cycles.st ---- *)
(* IEC 61131-3 §6.6.3.2 / Table 43 (TON), Table 44 (TOF), Table 45 (TP): TON.Q rises once IN has been TRUE for PT and falls with IN; TOF.Q holds for PT after IN falls; TP.Q is a single pulse of width PT regardless of IN. Time is the simulated clock advanced by the fixed cycle time (10 ms per cycle here), so elapsed time is exact. *)
FUNCTION_BLOCK TEST_TimersCycles
VAR
  ton : TON;
  tof : TOF;
  tp : TP;
  inp : BOOL;
  cycles : DINT;
END_VAR
METHOD Cycle
  ton(IN := inp, PT := T#50ms);
  tof(IN := inp, PT := T#50ms);
  tp(IN := inp, PT := T#30ms);
END_METHOD
METHOD Test_TonFiresAfterPreset
  inp := TRUE;
  RUN_CYCLES(4);
  ASSERT_FALSE(ton.Q);
  RUN_CYCLES(2);
  ASSERT_TRUE(ton.Q);
END_METHOD
METHOD Test_TonResetsWhenInputFalls
  inp := TRUE;
  RUN_CYCLES(10);
  ASSERT_TRUE(ton.Q);
  inp := FALSE;
  RUN_CYCLES(1);
  ASSERT_FALSE(ton.Q);
  ASSERT_EQUAL_TIME(ton.ET, T#0ms);
END_METHOD
METHOD Test_TonElapsedSaturatesAtPreset
  inp := TRUE;
  RUN_CYCLES(20);
  ASSERT_EQUAL_TIME(ton.ET, T#50ms);
END_METHOD
METHOD Test_TonShortPulseNeverFires
  inp := TRUE;
  RUN_CYCLES(3);
  inp := FALSE;
  RUN_CYCLES(1);
  inp := TRUE;
  RUN_CYCLES(3);
  ASSERT_FALSE(ton.Q);
END_METHOD
METHOD Test_TofHoldsAfterInputFalls
  inp := TRUE;
  RUN_CYCLES(2);
  ASSERT_TRUE(tof.Q);
  inp := FALSE;
  RUN_CYCLES(3);
  ASSERT_TRUE(tof.Q);
  RUN_CYCLES(4);
  ASSERT_FALSE(tof.Q);
END_METHOD
METHOD Test_TpPulseWidth
  inp := TRUE;
  RUN_CYCLES(1);
  ASSERT_TRUE(tp.Q);
  RUN_CYCLES(1);
  ASSERT_TRUE(tp.Q);
  RUN_CYCLES(5);
  ASSERT_FALSE(tp.Q);
END_METHOD
METHOD Test_TpIgnoresInputFallingMidPulse
  inp := TRUE;
  RUN_CYCLES(1);
  inp := FALSE;
  RUN_CYCLES(1);
  ASSERT_TRUE(tp.Q);
END_METHOD
METHOD Test_RunUntilReturnsCyclesToFire
  inp := TRUE;
  cycles := RUN_UNTIL('ton.Q', 100);
  ASSERT_EQUAL_DINT(cycles, 6);
END_METHOD
END_FUNCTION_BLOCK

(* ---- widening.st ---- *)
(* IEC 61131-3 §6.6.1 / Table 30 (ANY_NUM typing): in a mixed-type operation both operands widen to the wider type, so SINT+INT is INT, INT+DINT is DINT, DINT+REAL is REAL, REAL+LREAL is LREAL; the operation is evaluated at the wider type and does not wrap at the narrower one. *)
FUNCTION_BLOCK TEST_Widening
VAR s : SINT; i : INT; d : DINT; r : REAL; l : LREAL; u : USINT; END_VAR
METHOD Test_SintPlusIntIsInt
  s := 100; i := 1000;
  ASSERT_EQUAL_INT(s + i, 1100);
END_METHOD
METHOD Test_SintPlusSintWrapsAtSint
  s := 100;
  s := s + s;
  ASSERT_EQUAL_SINT(s, -56);
END_METHOD
METHOD Test_NoNarrowWrapInWiderExpression
  s := 100; i := 0;
  d := s + i + s;
  ASSERT_EQUAL_DINT(d, 200);
END_METHOD
METHOD Test_IntPlusDintIsDint
  i := 30000; d := 100000;
  ASSERT_EQUAL_DINT(i + d, 130000);
END_METHOD
METHOD Test_DintPlusRealIsReal
  d := 3; r := 0.5;
  ASSERT_EQUAL_REAL(d + r, 3.5);
END_METHOD
METHOD Test_RealPlusLrealIsLreal
  r := 1.5; l := 0.25;
  ASSERT_EQUAL_LREAL(r + l, 1.75);
END_METHOD
METHOD Test_IntTimesDint
  i := 20000; d := 2;
  ASSERT_EQUAL_DINT(i * d, 40000);
END_METHOD
METHOD Test_UsintPlusSintIsInt
  u := 200; s := -100;
  ASSERT_EQUAL_INT(u + s, 100);
END_METHOD
END_FUNCTION_BLOCK
